{attribute 'qualified_only'}
VAR_GLOBAL PERSISTENT
	stRecipe : ST_PersistentRecipe;
	arCal : ARRAY[1..3] OF ST_PersistentInner;
END_VAR
VAR_GLOBAL
	fbCell : FB_PersistentCell;
	aCells : ARRAY[1..2] OF FB_PersistentCell;
END_VAR

(* stored: Version 1.1.0.1
   GVL GVL_Persistent: Id {3f6a1c52-8d7e-4b0a-9a41-5c2e7d9b1a04} *)
